FUNCTION_BLOCK RawToEng
VAR_INPUT
	iEnabled : BOOL;
	wRawValue : WORD;
	AnalogConversion : TAnalogConversion;
END_VAR
VAR_OUTPUT
	oEnabled : BOOL;
	fScaledValue : REAL;
END_VAR
VAR
END_VAR

//Prepocet z wRawValue (z procesu po ModbusTCP) na fScaledValue (do PLC) podle parametru v AnalogConversion.

//Filtrace hodnoty: odfiltrovani skokoveho kmitani z minimalniho rozsahu na maximalni hodnotu >= 27648 (podteceni sumu u nuly v simulatoru)
IF wRawValue >= AnalogConversion.TransducerHiLevel THEN 
	IF fScaledValue < ((AnalogConversion.ScaledValHiLevel + AnalogConversion.ScaledValLoLevel) / 2.0) THEN
		wRawValue := AnalogConversion.TransducerLoLevel;
	ELSE
		wRawValue := AnalogConversion.TransducerHiLevel;
	END_IF;
END_IF;

fScaledValue := (AnalogConversion.ScaledValHiLevel - AnalogConversion.ScaledValLoLevel) * WORD_TO_REAL(wRawValue - AnalogConversion.TransducerLoLevel) / UINT_TO_REAL(AnalogConversion.TransducerHiLevel - AnalogConversion.TransducerLoLevel) + AnalogConversion.ScaledValLoLevel;
oEnabled := iEnabled;

END_FUNCTION_BLOCK

(* stored: Version 1.1.0.1, ProductVersion 3.1.4024.13
   POU RawToEng: Id {2bc2853a-1077-4f1d-a7fb-ade6d5b9212b}, SpecialFunc None *)
